{region 'Documentation'}
(*!
<summary>Checks the observed value sequence; Evaluate also checks the current value and
completeness.</summary>
<description>

Uses the whole Expected array from its declared lower bound. Keep its binding, bounds and
values stable until Reset; supply it on reset and disabled FB calls as well.

Observation accepts the current expected value and then permits advancing by one element
on a later change. Repeated equal values do not advance. An unexpected value or an out-of-range
sequence index reports Failed.

Evaluate checks the current value and requires the final expected element to have been
reached; only then can the result become Passed. Disabling observation retains progression.
Reset restarts it.

</description>
*)
{endregion}
FUNCTION_BLOCK AssertSequence_DInt EXTENDS AssertionWithEvaluationBase
VAR_INPUT
    IN : DINT; //! Actual value to observe.
END_VAR
VAR_IN_OUT CONSTANT
    Expected : ARRAY[*] OF DINT; //! Complete expected sequence; read without modifying the supplied array.
END_VAR
VAR
    FExpectedIndex : DINT;
    FSequenceIndexInitialized : BOOL;
    FAllowAdvance : BOOL;
END_VAR

SUPER^();

{region 'Documentation'}
(*!
<summary>Advances at most one entry and checks the current value before explicit completeness evaluation.</summary>
*)
{endregion}
METHOD PROTECTED Assert
VAR
    LowerIndex : DINT;
    UpperIndex : DINT;
    ExpectedValue : DINT;
    MatchesExpected : BOOL;
    AllowAdvance : BOOL;
    Message : STRING(GVL_Constants.MessageLength);
    ExpectedText : STRING(GVL_Constants.AssertionValueLength);
    ActualText : STRING(GVL_Constants.AssertionValueLength);
END_VAR
LowerIndex := LOWER_BOUND(Expected, 1);
UpperIndex := UPPER_BOUND(Expected, 1);

IF NOT FSequenceIndexInitialized THEN
    FExpectedIndex := LowerIndex;
    FSequenceIndexInitialized := TRUE;
END_IF;

IF NOT (ObservationActive OR EvaluationActive) THEN
    RETURN;
END_IF;

IF Result = E_Result.Error THEN
    RETURN;
END_IF;

IF Result = E_Result.Failed THEN
    RETURN;
END_IF;

IF (FExpectedIndex < LowerIndex) OR (FExpectedIndex > UpperIndex) THEN
    Message := CONCAT('Assertion failed: sequence index out of range. ExpectedIndex = ',
        DINT_TO_STRING(FExpectedIndex));
    Message := CONCAT(Message, ', LowerIndex = ');
    Message := CONCAT(Message, DINT_TO_STRING(LowerIndex));
    Message := CONCAT(Message, ', UpperIndex = ');
    Message := CONCAT(Message, DINT_TO_STRING(UpperIndex));
    Message := CONCAT(Message, '.');
    Fail(Message := Message);
    RETURN;
END_IF;

AllowAdvance := FAllowAdvance;
IF ObservationActive THEN
    FAllowAdvance := TRUE;
END_IF;

ExpectedValue := Expected[FExpectedIndex];
MatchesExpected := IN = ExpectedValue;

IF AllowAdvance AND NOT MatchesExpected THEN
    IF FExpectedIndex = UpperIndex THEN
        Message := CONCAT('Assertion failed: sequence continued beyond its last entry. LastIndex = ',
            DINT_TO_STRING(UpperIndex));
        Message := CONCAT(Message, '.');
        Fail(Message := Message);
        RETURN;
    END_IF;

    FExpectedIndex := FExpectedIndex + 1;
    ExpectedValue := Expected[FExpectedIndex];
    MatchesExpected := IN = ExpectedValue;
END_IF;

IF NOT MatchesExpected THEN
    ExpectedText := DINT_TO_STRING(ExpectedValue);
    ActualText := DINT_TO_STRING(IN);
    Message := CONCAT('Assertion failed: sequence value does not match. ExpectedIndex = ',
        DINT_TO_STRING(FExpectedIndex));
    Message := CONCAT(Message, ', Expected = ');
    Message := CONCAT(Message, ExpectedText);
    Message := CONCAT(Message, ', Actual = ');
    Message := CONCAT(Message, ActualText);
    Message := CONCAT(Message, '.');
    Fail(Message := Message);
    RETURN;
END_IF;

IF NOT EvaluationActive THEN
    RETURN;
END_IF;

IF FExpectedIndex <> UpperIndex THEN
    Message := CONCAT('Assertion failed: sequence is incomplete. ExpectedIndex = ',
        DINT_TO_STRING(FExpectedIndex));
    Message := CONCAT(Message, ', LastIndex = ');
    Message := CONCAT(Message, DINT_TO_STRING(UpperIndex));
    Message := CONCAT(Message, '.');
    Fail(Message := Message);
    RETURN;
END_IF;

Pass();
END_METHOD

{region 'Documentation'}
(*!
<summary>Restart progression at the bound Expected array's lower index.</summary>
<description>

Runs only during the reset FB call with Expected supplied, not directly from Reset or
Initialize. Clears permission to advance from a previous observation.

</description>
*)
{endregion}
METHOD PROTECTED ResetAssertion
FExpectedIndex := LOWER_BOUND(Expected, 1);
FSequenceIndexInitialized := TRUE;
FAllowAdvance := FALSE;
END_METHOD

END_FUNCTION_BLOCK

(* stored: Version 1.1.0.1
   POU AssertSequence_DInt: Id {07b582c4-4cd6-4601-aefc-863ee17d986b}, SpecialFunc None
   Folder Internal: Id {e33b2c37-aa92-40c6-902f-987d57422beb}
   Method Assert: Id {15867031-1773-4f1c-b7b3-a5a661b76c7a}
   Method ResetAssertion: Id {52f35d45-b905-4213-9275-b7818e2235b0} *)
